(* IEC 61131-3 sources: Test-Git_ESME26/TestProgettoESME_26.fbsproj/PacDriveLib Migration/Motion/Control, 3 files *)

(* ---- PDL_FB_Brake.fb.st ---- *)
FUNCTION_BLOCK PDL_FB_Brake
VAR_INPUT
	i_xEnable  : BOOL;
	i_xRelease : BOOL;
	i_ifDrive  : Moin.IF_Axis;
END_VAR
VAR_OUTPUT
	q_xActive   : BOOL;
	q_xReady    : BOOL;
	q_etDiag    : GD.ET_Diag     := GD.ET_Diag.Ok;
	q_etDiagExt : PDL_ET_DiagExt := PDL_ET_DiagExt.Disabled;
	q_sMsg      : STRING[80];
	q_xReleased : BOOL;
END_VAR
VAR
	xSuccess                 : BOOL;
	ifDeviceTreeObjectAccess : UFMPLCI.IF_DeviceTreeObjectAccess;
	sDriveName               : STRING(80);
	ifBrakeAccess            : DDI.IF_BrakeAccess;
	ifBrake                  : DDI.IF_Brake;
	ifGetParentDevice        : DTSI.IF_GetParentDevice;
	ifDeviceAccess           : DTSI.IF_DeviceAccess;
	ifWorkingModeAccess      : CFDI.IF_WorkingModeAccess;
	ifWorkingMode            : CFDI.IF_WorkingMode;
	etWorkingState           : CFDI.ET_WorkingState;
	etSercosState            : SMI.ET_SercosState;
	etAxisState              : MOIN.ET_AxisState;
	etDiagExt                : PDL_ET_DiagExt := PDL_ET_DiagExt.Disabled;
	diState                  : DINT;
	xEnableFlag              : BOOL;
	fbLoggerPoint            : APL.FB_LoggerPoint;
	fbBrakeReleaseSet        : FB_BrakeReleaseSet;
	fbBrakeDisconnectionTime : FB_BrakeDisconnectionTime;
	fbBrakeCouplingTime      : FB_BrakeCouplingTime;
	xError                   : BOOL;
	tonTimeOutBrake          : Standard.TON;
	tonTimeOutException      : Standard.TON;
	tBrakeCouplingTemp       : TIME := T#500MS;
	tBrakeDisconnectTemp     : TIME := T#500MS;
	sResultMsg               : STRING(80);
	etResult                 : SE_Async.ET_Result;

END_VAR
VAR CONSTANT
	c_timTimeOutException : TIME := T#1S;
END_VAR

IF i_xEnable AND NOT xEnableFlag THEN (* Input action *)
	xEnableFlag := TRUE;

	THIS^.fbLoggerPoint.AddLogEntry(
		i_etLogLevel := APL.ET_LogLevel.UserAction,
		i_etDiag     := q_etDiag,
		i_udiDiagExt := q_etDiagExt,
		i_sMessage   := 'enable function block',
		q_etDiag     =>,
		q_etDiagExt  => );

	q_xActive   := TRUE;
	q_xReady    := FALSE;
	q_xReleased := FALSE;
	SetDiagOutput(
		i_etDiag    := GD.ET_Diag.Ok,
		i_etDiagExt := PDL_ET_DiagExt.Initializing,
		i_sMsg      := '');
	xSuccess := InitInterfaces();
	IF NOT xSuccess THEN
		RETURN;
	ELSE
		IF SE_Async.G_ifAsyncMgr.xInitDone THEN
			q_xReady    := TRUE;
			q_xReleased := (ifBrake.BrakeState = DDI.ET_BrakeState.released);
			IF q_xReleased THEN // Bremse is open --> wait for closing Brake (i_xRelease = false)
				SetDiagOutput(
					i_etDiag    := GD.ET_Diag.Ok,
					i_etDiagExt := PDL_ET_DiagExt.WaitForNotRelease,
					i_sMsg      := '');
				diState := 40;
			ELSE // brake is closed --> wait for opening brake (i_xRelease = true)
				SetDiagOutput(
					i_etDiag    := GD.ET_Diag.Ok,
					i_etDiagExt := PDL_ET_DiagExt.WaitForRelease,
					i_sMsg      := '');
				diState := 10;
			END_IF
		ELSE
			SE_Async.G_ifAsyncMgr.Init();
			diState := 150;
		END_IF
	END_IF

ELSIF NOT i_xEnable AND xEnableFlag AND q_xActive THEN
	xEnableFlag := FALSE;
	THIS^.fbLoggerPoint.AddLogEntry(
		i_etLogLevel := APL.ET_LogLevel.UserAction,
		i_etDiag     := q_etDiag,
		i_udiDiagExt := q_etDiagExt,
		i_sMessage   := 'disable function block',
		q_etDiag     =>,
		q_etDiagExt  => );
	SetDiagOutput(
		i_etDiag    := GD.ET_Diag.Ok,
		i_etDiagExt := PDL_ET_DiagExt.WaitUntilDisabled,
		i_sMsg      := '');

	q_xReady := FALSE;
	IF diState = 10 THEN // Brake is already closed
		diState := 120;
	ELSE
		fbBrakeReleaseSet.ifBrake  := ifBrake;
		fbBrakeReleaseSet.xRelease := FALSE;
		SE_Async.G_ifAsyncMgr.Start(
			i_ifAsync    := fbBrakeReleaseSet,
			q_etResult   => etResult,
			q_sResultMsg => sResultMsg,
			q_xError     => xError);
		IF xError THEN
			diState := 120;
		ELSE
			tonTimeOutBrake(IN := FALSE, PT := c_timTimeOutException);
			diState := 100;
		END_IF
	END_IF
END_IF

IF q_xReady THEN
	etSercosState  := FC_GetSercosState();
	etWorkingState := ifWorkingMode.ActualState;
	etAxisState    := i_ifDrive.etAxisState;
	IF etSercosState <> SMI.ET_SercosState.Phase4 THEN
		q_xReady    := FALSE;
		q_xReleased := FALSE;
		SetDiagOutput(
			i_etDiag    := GD.ET_Diag.SercosConditionInvalid,
			i_etDiagExt := PDL_ET_DiagExt.SercosNotInPhaseFour,
			i_sMsg      := 'Sercos not in phase four');
		diState := 0;
	ELSIF etWorkingState = CFDI.ET_WorkingState.Deactivated THEN
		q_xReady    := FALSE;
		q_xReleased := FALSE;
		SetDiagOutput(
			i_etDiag    := GD.ET_Diag.DriveConditionInvalid,
			i_etDiagExt := PDL_ET_DiagExt.DriveNotReady,
			i_sMsg		:= STANDARD.CONCAT(sDriveName, '.WorkingMode = deactivated'));
		diState := 0;
	ELSIF etAxisState <> Moin.ET_AxisState.Disabled THEN
		q_xReady    := FALSE;
		q_xReleased := FALSE;
		SetDiagOutput(
			i_etDiag    := GD.ET_Diag.DriveConditionInvalid,
			i_etDiagExt := PDL_ET_DiagExt.DriveNotReady,
			i_sMsg		:= STANDARD.CONCAT(sDriveName, '.AxisState <> Disabled; Drive has to be disabled'));
		diState := 0;
	END_IF
END_IF

CASE diState OF
	0: (* No operation / FB disabled *)
		;
	10: // Brake closed, wait for releasing Brake (i_xRelease = true)
		IF i_xRelease THEN // input release Brake
			fbLoggerPoint.AddLogEntry(
				i_etLogLevel := APL.ET_LogLevel.UserAction,
				i_etDiag     := q_etDiag,
				i_udiDiagExt := q_etDiagExt,
				i_sMessage   := 'Release Brake - read out disconnection time',
				q_etDiag     =>,
				q_etDiagExt  => );
			etSercosState := FC_GetSercosState();
			fbBrakeDisconnectionTime.ifBrake  := ifBrake;
			SE_Async.G_ifAsyncMgr.Start(
				i_ifAsync    := fbBrakeDisconnectionTime, // read Disconnecting time from Drive
				q_etResult   => etResult,
				q_sResultMsg => sResultMsg,
				q_xError     => xError);
			IF xError THEN
				IF etResult = SE_Async.ET_Result.MaxNumOfReusableObjectsExceeded THEN
					diState := diState; // Try again to Start Async in next cycle
				ELSE
					AsyncExtDiagTranslation();
					diState := 200;
				END_IF
			ELSE
				tonTimeOutBrake(IN := FALSE, PT := c_timTimeOutException);
				diState := 15;
			END_IF
		END_IF
	15: // Wait for BrakeDisconnectionTime has been read
		tonTimeOutBrake(IN := TRUE);
		IF fbBrakeDisconnectionTime.xDone THEN
			tBrakeDisconnectTemp       := fbBrakeDisconnectionTime.timTime;
			fbBrakeReleaseSet.ifBrake  := ifBrake;
			fbBrakeReleaseSet.xRelease := TRUE;
			SE_Async.G_ifAsyncMgr.Start(
				i_ifAsync    := fbBrakeReleaseSet,
				q_etResult   => etResult,
				q_sResultMsg => sResultMsg,
				q_xError     => xError);
			IF xError THEN
				IF etResult = SE_Async.ET_Result.MaxNumOfReusableObjectsExceeded THEN
					diState := diState; // Try again to Start Async in next cycle
				ELSE
					AsyncExtDiagTranslation();
					diState := 200;
				END_IF
			ELSE
				fbLoggerPoint.AddLogEntry(
					i_etLogLevel := APL.ET_LogLevel.DebugMessage,
					i_etDiag     := q_etDiag,
					i_udiDiagExt := q_etDiagExt,
					i_sMessage   := 'Release Brake - brake release set',
					q_etDiag     =>,
					q_etDiagExt  => );
				tonTimeOutBrake(IN := FALSE, PT := c_timTimeOutException);
				diState := 20;
			END_IF
		ELSIF tonTimeOutBrake.Q THEN
			SetDiagOutput(
				i_etDiag    := GD.ET_Diag.UnexpectedProgramBehavior,
				i_etDiagExt := PDL_ET_DiagExt.AsyncAddWasNotSuccessful,
				i_sMsg      := 'Timeout at read of BrakeDisconnectionTime');
			diState := 200;
		END_IF
	20: // Wait for Brake is release, Release Commando Done
		tonTimeOutBrake(IN := TRUE);
		IF fbBrakeReleaseSet.xDone THEN
			SetDiagOutput(
				i_etDiag    := GD.ET_Diag.Ok,
				i_etDiagExt := PDL_ET_DiagExt.WaitUntilBrakeReleased,
				i_sMsg      := '');
			tonTimeOutBrake(IN := FALSE, PT := tBrakeDisconnectTemp);
			tonTimeOutException(IN := FALSE, PT := c_timTimeOutException);
			diState := 25;
		ELSIF tonTimeOutBrake.Q THEN
			SetDiagOutput(
				i_etDiag    := GD.ET_Diag.UnexpectedProgramBehavior,
				i_etDiagExt := PDL_ET_DiagExt.AsyncAddWasNotSuccessful,
				i_sMsg      := 'Timeout at BrakeReleaseSet');
			diState := 200;
		END_IF
	25: // wait till brake has to be open (check both, system signal and own time out)
		tonTimeOutBrake(IN := TRUE);
		tonTimeOutException(IN := TRUE);
		IF tonTimeOutBrake.Q THEN
			IF (ifBrake.BrakeState = DDI.ET_BrakeState.released) THEN // Brake is released
				q_xReleased := TRUE;
				SetDiagOutput(
					i_etDiag    := GD.ET_Diag.Ok,
					i_etDiagExt := PDL_ET_DiagExt.WaitForNotRelease,
					i_sMsg      := '');
				diState := 40;
			ELSE
				SetDiagOutput(
					i_etDiag    := GD.ET_Diag.UnexpectedProgramBehavior,
					i_etDiagExt := PDL_ET_DiagExt.BrakeStateChangedNotInTime,
					i_sMsg      := 'Timeout at wait for Brake Release');
				diState := 200;
			END_IF
		ELSIF tonTimeOutException.Q THEN
			SetDiagOutput(
				i_etDiag    := GD.ET_Diag.UnexpectedProgramBehavior,
				i_etDiagExt := PDL_ET_DiagExt.BrakeStateChangedNotInTime,
				i_sMsg      := 'Timeout at wait for Brake Release');
			diState := 200;
		END_IF
	40: // Brake released, wait for Brake is coupled (i_xRelease = FALSE)
		IF NOT i_xRelease THEN
			fbLoggerPoint.AddLogEntry(
				i_etLogLevel := APL.ET_LogLevel.UserAction,
				i_etDiag     := q_etDiag,
				i_udiDiagExt := q_etDiagExt,
				i_sMessage   := 'Close Brake - read out coupling time',
				q_etDiag     =>,
				q_etDiagExt  => );
			fbBrakeCouplingTime.ifBrake  := ifBrake;
			SE_Async.G_ifAsyncMgr.Start(
				i_ifAsync    := fbBrakeCouplingTime,
				q_etResult   => etResult,
				q_sResultMsg => sResultMsg,
				q_xError     => xError);
			IF xError THEN
				IF etResult = SE_Async.ET_Result.MaxNumOfReusableObjectsExceeded THEN
					diState := diState; // Try again to Start Async in next cycle
				ELSE
					AsyncExtDiagTranslation();
					diState := 200;
				END_IF
			ELSE
				tonTimeOutBrake(IN := FALSE, PT := c_timTimeOutException);
				diState := 45;
			END_IF
		END_IF
	45: // wait for BrakeCouplingTime has been read out
		tonTimeOutBrake(IN := TRUE);
		IF fbBrakeCouplingTime.xDone THEN
			tBrakeCouplingTemp         := fbBrakeCouplingTime.timTime;
			fbBrakeReleaseSet.ifBrake  := ifBrake;
			fbBrakeReleaseSet.xRelease := FALSE;
			SE_Async.G_ifAsyncMgr.Start(
				i_ifAsync    := fbBrakeReleaseSet,
				q_etResult   => etResult,
				q_sResultMsg => sResultMsg,
				q_xError     => xError);
			IF xError THEN
				AsyncExtDiagTranslation();
				diState := 200;
			ELSE
				fbLoggerPoint.AddLogEntry(
					i_etLogLevel := APL.ET_LogLevel.DebugMessage,
					i_etDiag     := q_etDiag,
					i_udiDiagExt := q_etDiagExt,
					i_sMessage   := 'Close Brake - brake release set',
					q_etDiag     =>,
					q_etDiagExt  => );
				tonTimeOutBrake(IN := FALSE, PT := c_timTimeOutException);
				diState := 50;
			END_IF
		ELSIF tonTimeOutBrake.Q THEN
			SetDiagOutput(
				i_etDiag    := GD.ET_Diag.UnexpectedProgramBehavior,
				i_etDiagExt := PDL_ET_DiagExt.AsyncAddWasNotSuccessful,
				i_sMsg      := 'Timeout at read of BrakeCouplingTime');
			diState := 200;
		END_IF
	50: // Wait for BrakeRelaseSet Done
		tonTimeOutBrake(IN := TRUE);
		IF fbBrakeReleaseSet.xDone THEN
			SetDiagOutput(
				i_etDiag    := GD.ET_Diag.Ok,
				i_etDiagExt := PDL_ET_DiagExt.WaitUntilBrakeClosed,
				i_sMsg      := '');
			tonTimeOutBrake(IN := FALSE, PT := tBrakeCouplingTemp);
			tonTimeOutException(IN := FALSE, PT := c_timTimeOutException);
			diState := 55;
		ELSIF tonTimeOutBrake.Q THEN
			SetDiagOutput(
				i_etDiag    := GD.ET_Diag.UnexpectedProgramBehavior,
				i_etDiagExt := PDL_ET_DiagExt.AsyncAddWasNotSuccessful,
				i_sMsg      := 'Timeout at BrakeReleaseSet');
			diState := 200;
		END_IF
	55: // wait till brake is closed (check both, system signal and own time out)
		tonTimeOutBrake(IN := TRUE);
		tonTimeOutException(IN := TRUE);
		IF tonTimeOutBrake.Q THEN
			IF (ifBrake.BrakeState = DDI.ET_BrakeState.coupled)  THEN
				tonTimeOutException(IN := FALSE);
				tonTimeOutBrake(IN := FALSE);
				q_xReleased := FALSE;
				SetDiagOutput(
					i_etDiag    := GD.ET_Diag.Ok,
					i_etDiagExt := PDL_ET_DiagExt.WaitForRelease,
					i_sMsg      := '');
				diState := 10;
			ELSE
				SetDiagOutput(
					i_etDiag    := GD.ET_Diag.UnexpectedProgramBehavior,
					i_etDiagExt := PDL_ET_DiagExt.BrakeStateChangedNotInTime,
					i_sMsg      := 'Timeout at wait for Brake coupled');
				diState := 200;
			END_IF
		ELSIF tonTimeOutBrake.Q THEN
			SetDiagOutput(
				i_etDiag    := GD.ET_Diag.UnexpectedProgramBehavior,
				i_etDiagExt := PDL_ET_DiagExt.BrakeStateChangedNotInTime,
				i_sMsg      := 'Timeout at wait for Brake Close');
			diState := 200;
		END_IF

		//---------------------------------------------------------------------------------
	100:
		tonTimeOutBrake(IN := TRUE);
		IF fbBrakeReleaseSet.xDone THEN
			IF i_ifDrive.etAxisState = MOIN.ET_AxisState.Disabled THEN
				tonTimeOutBrake(IN := FALSE, PT := c_timTimeOutException);
				diState := 110;
			ELSE
				diState := 120;
			END_IF
		ELSIF tonTimeOutBrake.Q THEN
			SetDiagOutput(
				i_etDiag    := GD.ET_Diag.UnexpectedProgramBehavior,
				i_etDiagExt := PDL_ET_DiagExt.AsyncAddWasNotSuccessful,
				i_sMsg      := 'Timeout at FC_BrakeReleaseSet');
			diState := 120;
		END_IF
	110: (* AxisState = 1 or 2 *)
		tonTimeOutBrake(IN := TRUE);
		IF (ifBrake.BrakeState = DDI.ET_BrakeState.coupled) THEN
			tonTimeOutBrake(IN := FALSE, PT := tBrakeCouplingTemp);
			diState := 115;
		ELSIF tonTimeOutBrake.Q THEN
			SetDiagOutput(
				i_etDiag    := GD.ET_Diag.UnexpectedProgramBehavior,
				i_etDiagExt := PDL_ET_DiagExt.BrakeStateChangedNotInTime,
				i_sMsg      := 'Timeout at wait for Brake Close');
			diState := 120;
		END_IF
	115:
		tonTimeOutBrake(IN := TRUE);
		IF tonTimeOutBrake.Q THEN
			diState := 120;
		END_IF
	120:
		q_xActive   := FALSE;
		q_xReady    := FALSE;
		q_xReleased := FALSE;
		SetDiagOutput(
			i_etDiag    := GD.ET_Diag.Ok,
			i_etDiagExt := PDL_ET_DiagExt.Disabled,
			i_sMsg      := '');
		tonTimeOutBrake(IN := FALSE);
		diState := 0;

	150:
		SE_Async.G_ifAsyncMgr.Init(
			q_xError     => xError,
			q_etResult   => etResult,
			q_sResultMsg => sResultMsg);
		IF xError THEN
			AsyncExtDiagTranslation();
			diState := 200;
		ELSIF SE_Async.G_ifAsyncMgr.xInitDone THEN
			q_xReady    := TRUE;
			q_xReleased := (ifBrake.BrakeState = DDI.ET_BrakeState.released);
			IF q_xReleased THEN // Bremse is open --> wait for closing Brake (i_xRelease = false)
				SetDiagOutput(
					i_etDiag    := GD.ET_Diag.Ok,
					i_etDiagExt := PDL_ET_DiagExt.WaitForNotRelease,
					i_sMsg      := '');
				diState := 40;
			ELSE // brake is closed --> wait for opening brake (i_xRelease = true)
				SetDiagOutput(
					i_etDiag    := GD.ET_Diag.Ok,
					i_etDiagExt := PDL_ET_DiagExt.WaitForRelease,
					i_sMsg      := '');
				diState := 10;
			END_IF
		END_IF

	200:
		q_xReady    := FALSE;
		q_xReleased := (ifBrake.BrakeState = DDI.ET_BrakeState.released);
		diState := 0;

END_CASE

(* ---- PDL_FB_DriveEnable.fb.st ---- *)
FUNCTION_BLOCK PDL_FB_DriveEnable
VAR_INPUT
	i_xEnable      : BOOL; (* Enable of FB *)
	i_ifDrive      : MOIN.IF_Axis; (* Axis *)
	i_xEnableDrive : BOOL; (* Power on *)
	i_xDiagQuit    : BOOL; (* reset error *)
END_VAR

VAR_OUTPUT
	q_xActive       : BOOL; (* FB enabled*)
	q_xReady        : BOOL;
	q_etDiag        : GD.ET_Diag     := GD.ET_Diag.Ok;
	q_etDiagExt     : PDL_ET_DiagExt := PDL_ET_DiagExt.Disabled;
	q_sMsg          : STRING[80];
	q_xDriveEnabled : BOOL; (* power is on*)
END_VAR

VAR
	xInterfacesInitialised : BOOL;

	xEnableFlag : BOOL;
	diState     : DINT;

	rtrigDiagQuit    : Standard.R_TRIG;
	xDriveEnabledOld : BOOL;

	fbLoggerPoint : APL.FB_LoggerPoint;

	fbPower : PLCO.MC_Power;
	fbStop  : PLCO.MC_Stop;
	fbReset	: PLCO.MC_Reset;

	ifDeviceTreeObjectAccess      : UFMPLCI.IF_DeviceTreeObjectAccess;
	sDriveName                    : STRING(80);
	ifGetParentDevice             : DTSI.IF_GetParentDevice;
	ifDiagnostic                  : UFMPLCI.IF_Diagnostic;
	ifDiagnosticAccess            : UFMPLCI.IF_DiagnosticAccess;
	ifDeviceAccess                : DTSI.IF_DeviceAccess;
	ifPowerSupply                 : DDI.IF_PowerSupply;
	ifPowerSupplyAccess           : DDI.IF_PowerSupplyAccess;
	ifDrivePowerSupply            : DDI.IF_DrivePowerSupply;
	ifDrivePowerSupplyAccess      : DDI.IF_DrivePowerSupplyAccess;
	ifDriveConfigAccess           : DDI.IF_DriveConfigAccess;
	ifDriveConfig                 : DDI.IF_DriveConfig;
	ifWorkingModeAccess           : CFDI.IF_WorkingModeAccess;
	ifWorkingMode                 : CFDI.IF_WorkingMode;
	ifPowerSupplyDiagnosticAccess : UFMPLCI.IF_DiagnosticAccess;
	ifPowerSupplyDiagnostic       : UFMPLCI.IF_Diagnostic;
	ifPowerSupplyDevice           : DDI.DeviceTypeInterfaces.IF_Device_Type;
	xSuccess                      : BOOL;
	etSercosState                 : SMI.ET_SercosState;
	tonTimeOut                    : Standard.TON;
	xDriveIsReal                  : BOOL;
END_VAR
VAR CONSTANT
	c_timTimeoutPowerSupplyReady  : TIME := T#2000MS;
	c_timTimeoutPowerSupplyEnable : TIME := T#2000MS;
END_VAR

(*--------------------------------------------------------------------------------------------------------------------------------------------*)
//Enable
{region "enable"}
IF i_xEnable AND NOT xEnableFlag THEN
	xEnableFlag := TRUE;

	THIS^.fbLoggerPoint.AddLogEntry(	i_etLogLevel	:= APL.ET_LogLevel.UserAction,
										i_etDiag		:= q_etDiag,
										i_udiDiagExt	:= q_etDiagExt,
										i_sMessage		:= 'enable function block',
										q_etDiag		=> ,
										q_etDiagExt		=> );
	q_xActive			:= TRUE;
	q_xDriveEnabled		:= FALSE;

	IF NOT Init() THEN
		q_xReady			    := FALSE;
		xInterfacesInitialised  := FALSE;
		diState := 200;
	ELSE
		q_xReady 				:= TRUE;
		xInterfacesInitialised  := TRUE;
		SetDiagOutput(	i_etDiag	:= GD.ET_Diag.Ok,
						i_etDiagExt := PDL_ET_DiagExt.WaitForEnableDrive,
						i_sMsg		:= '');
		diState	:= 10;
	END_IF
{endregion}

(*--------------------------------------------------------------------------------------------------------------------------------------------*)
//Disable
{region "disable"}
ELSIF NOT i_xEnable AND xEnableFlag THEN
	xEnableFlag := FALSE;
	THIS^.fbLoggerPoint.AddLogEntry(	i_etLogLevel	:= APL.ET_LogLevel.UserAction,
										i_etDiag		:= q_etDiag,
										i_udiDiagExt	:= q_etDiagExt,
										i_sMessage		:= 'disable function block',
										q_etDiag		=> ,
										q_etDiagExt		=> );
	q_xReady			:= FALSE;
	IF xInterfacesInitialised THEN
		SetDiagOutput(	i_etDiag	:= GD.ET_Diag.Ok,
						i_etDiagExt := PDL_ET_DiagExt.WaitUntilDriveDisabled,
						i_sMsg		:= '');

		diState := 100; // whait till axis disabled
	ELSE
		q_xActive			:= FALSE;
		q_xDriveEnabled		:= FALSE;

		SetDiagOutput(	i_etDiag	:= GD.ET_Diag.Ok,
						i_etDiagExt := PDL_ET_DiagExt.Disabled,
						i_sMsg		:= '');
		diState	:= 0;
	END_IF
END_IF
{endregion}

(*--------------------------------------------------------------------------------------------------------------------------------------------*)
// Cyclic when enabled
{region "cyclic"}
IF xInterfacesInitialised AND q_xActive THEN
	q_xDriveEnabled :=  i_ifDrive.etAxisState >= MOIN.ET_AxisState.Standstill;
	etSercosState := FC_GetSercosState();
	fbReset( Execute := FALSE );

	IF xDriveIsReal AND_THEN ifPowerSupplyDiagnostic.DiagClass >= 3 THEN
		fbPower( Enable := FALSE );
		q_xReady	:= FALSE;
		SetDiagOutput(	i_etDiag	:= GD.ET_Diag.PowerSupplyConditionInvalid,
						i_etDiagExt := PDL_ET_DiagExt.PowerSupplyNotReady,
						i_sMsg		:= SE_CTBX.FC_MultiConcat(	i_sString1 := 'DiagCode: ',
														i_sString2 := TO_STRING(ifPowerSupplyDiagnostic.DiagCode),
														i_sString3 := ' - DiagMsg: ',
														i_sString4 := ifPowerSupplyDiagnostic.DiagMsg));
		diState := 200;

	//check for drive errors
	ELSIF ifDiagnostic.DiagClass >= 3 THEN
		fbPower( Enable := FALSE );
		q_xReady		:= FALSE;
		q_xDriveEnabled := FALSE;
		SetDiagOutput(	i_etDiag	:= GD.ET_Diag.DriveConditionInvalid,
						i_etDiagExt := PDL_ET_DiagExt.DriveNotReady,
						i_sMsg		:= SE_CTBX.FC_MultiConcat(	i_sString1 := 'DiagCode: ',
																i_sString2 := TO_STRING(ifDiagnostic.DiagCode),
																i_sString3 := ' - DiagMsg: ',
																i_sString4 := ifDiagnostic.DiagMsg));
		diState := 200;

	//check sercos state
	ELSIF etSercosState <> SMI.ET_SercosState.Phase4 THEN
		fbPower( Enable := FALSE );
		q_xReady:= FALSE;
		q_xDriveEnabled:= FALSE;
		SetDiagOutput(	i_etDiag	:= GD.ET_Diag.SercosConditionInvalid,
						i_etDiagExt := PDL_ET_DiagExt.SercosNotInPhaseFour,
						i_sMsg		:= 'Sercos not in phase four');
		diState:= 200;

	//check inverter enable
	ELSIF xDriveIsReal AND_THEN NOT ifDrivePowerSupply.InverterEnable AND i_xEnableDrive THEN
		fbPower( Enable := FALSE );
		q_xReady			:= FALSE;
		q_xDriveEnabled		:= FALSE;
		SetDiagOutput(	i_etDiag	:= GD.ET_Diag.DriveConditionInvalid,
						i_etDiagExt := PDL_ET_DiagExt.InverterEnableOff,
						i_sMsg		:= sDriveName);
		diState := 200;
	END_IF

	//stop/disable drive
	IF    NOT i_xEnableDrive
	  AND diState = 10
	  AND fbPower.Enable
	THEN
		THIS^.fbLoggerPoint.AddLogEntry(	i_etLogLevel	:= APL.ET_LogLevel.UserAction,
											i_etDiag		:= q_etDiag,
											i_udiDiagExt	:= q_etDiagExt,
											i_sMessage		:= 'disable drive',
											q_etDiag		=> ,
											q_etDiagExt		=> );

		SetDiagOutput(	i_etDiag	:= GD.ET_Diag.Ok,
						i_etDiagExt := PDL_ET_DiagExt.WaitUntilDriveDisabled,
						i_sMsg		:= '');

		//if power on -> stop first
		IF fbPower.Status THEN
			diState := 30;
		ELSE
			diState := 100;
		END_IF
	END_IF

END_IF

IF q_xActive THEN
	rtrigDiagQuit(CLK := i_xDiagQuit);
END_IF
{endregion}

(*--------------------------------------------------------------------------------------------------------------------------------------------*)
//state machine
CASE diState OF

(*********************************************************************************************************************)
	0:	//Error or Not Enabled
		;

(*********************************************************************************************************************)
	10:	//enable drive
{region "enableDrive"}
		fbStop(Axis := i_ifDrive, Execute := FALSE );

		//set diag outpupt after enable cmd
		IF 	  i_xEnableDrive
		  AND NOT fbPower.Enable
		  AND i_xEnable
		THEN
			IF xDriveIsReal AND_THEN NOT ifPowerSupply.PowerSupplyCheck THEN
				ifPowerSupply.PowerSupplyCheckSet	:= TRUE;
				SetDiagOutput(	i_etDiag	:= GD.ET_Diag.Ok,
								i_etDiagExt := PDL_ET_DiagExt.WaitUntilPowerSupplyReady,
								i_sMsg		:= '');
				tonTimeout(IN := FALSE, PT := c_timTimeoutPowerSupplyReady);		(* init Timeout for PS Ready *)
				diState	:= 20;
				RETURN;
			ELSE
				THIS^.fbLoggerPoint.AddLogEntry(	i_etLogLevel	:= APL.ET_LogLevel.UserAction,
													i_etDiag		:= q_etDiag,
													i_udiDiagExt	:= q_etDiagExt,
													i_sMessage		:= 'enable drive',
													q_etDiag		=> ,
													q_etDiagExt		=> );

				SetDiagOutput(	i_etDiag	:= GD.ET_Diag.Ok,
								i_etDiagExt := PDL_ET_DiagExt.WaitUntilDriveEnabled,
								i_sMsg		:= '');
			END_IF
		END_IF

		//cmd power on
		fbPower( Enable :=  i_xEnableDrive AND i_xEnable );
		q_xDriveEnabled :=  i_ifDrive.etAxisState >= MOIN.ET_AxisState.Standstill;

		//set diag output when on
		IF    q_xDriveEnabled
		  AND NOT xDriveEnabledOld
		THEN
			SetDiagOutput(	i_etDiag	:= GD.ET_Diag.Ok,
							i_etDiagExt := PDL_ET_DiagExt.DriveEnabled,
							i_sMsg		:= '');
		END_IF

		//error
		IF fbPower.Error THEN
			q_xReady		:= FALSE;
			q_xDriveEnabled	:= FALSE;

			SetDiagOutput(	i_etDiag	:= GD.ET_Diag.UnexpectedProgramBehavior,
							i_etDiagExt := PDL_ET_DiagExt.UnexpectedFeedback,
							i_sMsg		:= CONCAT('MC_Power.ErrorID: ', PLCO.FC_EtResultToString( fbPower.ErrorID ) ));

			fbPower( Enable := FALSE );
			diState	:= 200;
		END_IF
{endregion}

(*********************************************************************************************************************)
	20: (* Wait for PowerSupply GroupState >= 2 *)
{region "error"}
		tonTimeout(IN := TRUE);
		IF ifPowerSupply.GroupState >= 2  THEN								(* GroupState on PS *)
			tonTimeout(IN := FALSE, PT := c_timTimeoutPowerSupplyEnable);	(* init Timeout for PS Enabled *)
			diState := 10;

		ELSIF tonTimeout.Q THEN
			q_xReady	:= FALSE;
			SetDiagOutput(	i_etDiag	:= GD.ET_Diag.PowerSupplyConditionInvalid,
							i_etDiagExt := PDL_ET_DiagExt.PowerSupplyNotReady,
							i_sMsg		:= SE_CTBX.FC_MultiConcat(	i_sString1 := 'DiagCode: ',
																	i_sString2 := TO_STRING(ifPowerSupplyDiagnostic.DiagCode),
																	i_sString3 := ' - DiagMsg: ',
																	i_sString4 := ifPowerSupplyDiagnostic.DiagMsg));
			diState := 10;
		END_IF
{endregion}

(*********************************************************************************************************************)
	30: //controllerStop
{region "controllerStop"}
		IF 	  i_ifDrive.etAxisState <> MOIN.ET_AxisState.Disabled
		  AND i_ifDrive.etAxisState <> MOIN.ET_AxisState.ErrorStop
		  AND i_ifDrive.etAxisState <> MOIN.ET_AxisState.Standstill
		  AND i_ifDrive.etAxisState <> MOIN.ET_AxisState.Stopping
		THEN
			fbStop.Execute 			:= TRUE;
			fbStop.Deceleration 	:= i_ifDrive.lrErrorStopDec;
			fbStop.Jerk 			:= i_ifDrive.lrErrorStopJerk;
		END_IF

		fbStop();

		//stopping done
		IF 	  i_ifDrive.etAxisState = MOIN.ET_AxisState.Disabled
		  OR  i_ifDrive.etAxisState = MOIN.ET_AxisState.ErrorStop
		  OR  i_ifDrive.etAxisState = MOIN.ET_AxisState.Standstill
		  OR  fbStop.Done
		THEN
			fbStop( Axis := i_ifDrive, Execute := FALSE );

			diState := 100;
		END_IF

		//error
		IF fbStop.Error AND fbStop.ErrorId <> PLCO.ET_Result.StoppingInterrupted THEN
			q_xReady		:= FALSE;
			q_xDriveEnabled	:= FALSE;

			fbStop( Axis := i_ifDrive, Execute := FALSE );
			SetDiagOutput(	i_etDiag	:= GD.ET_Diag.UnexpectedProgramBehavior,
							i_etDiagExt := PDL_ET_DiagExt.UnexpectedFeedback,
							i_sMsg		:= CONCAT('MC_Stop.ErrorID: ', PLCO.FC_EtResultToString(fbStop.ErrorID) ));
			diState := 100;
		END_IF
{endregion}

(*********************************************************************************************************************)
	100: //disable drive
{region "disableDrive"}
		fbStop( Execute := FALSE );
		fbPower( Enable :=  FALSE );

		q_xDriveEnabled := i_ifDrive.etAxisState >= MOIN.ET_AxisState.Standstill;

		//wait for power off
		IF NOT q_xDriveEnabled THEN
			IF NOT i_xEnable THEN
				q_xActive := FALSE;
				SetDiagOutput(	i_etDiag	:= GD.ET_Diag.Ok,
								i_etDiagExt := PDL_ET_DiagExt.Disabled,
								i_sMsg		:= '');
				diState	:= 0;
			ELSE
				SetDiagOutput(	i_etDiag	:= GD.ET_Diag.Ok,
								i_etDiagExt := PDL_ET_DiagExt.WaitForEnableDrive,
								i_sMsg		:= '');
				diState	:= 10;
			END_IF
		END_IF

		//error
		IF fbPower.Error THEN
			q_xReady		:= FALSE;
			q_xDriveEnabled	:= FALSE;

			SetDiagOutput(	i_etDiag	:= GD.ET_Diag.UnexpectedProgramBehavior,
							i_etDiagExt := PDL_ET_DiagExt.UnexpectedFeedback,
							i_sMsg		:= CONCAT('MC_Power.ErrorID: ', PLCO.FC_EtResultToString( fbPower.ErrorID ) ));
			fbStop( Execute := FALSE );
		  	IF i_xEnable THEN
				diState	:= 200;
			ELSE
				diState	:= 0;
			END_IF
		END_IF
{endregion}

(*********************************************************************************************************************)
	200: //error
{region "error"}
		IF rtrigDiagQuit.Q //wait for cmd diag quit
		THEN
			THIS^.fbLoggerPoint.AddLogEntry(	i_etLogLevel	:= APL.ET_LogLevel.UserAction,
												i_etDiag		:= q_etDiag,
												i_udiDiagExt	:= q_etDiagExt,
												i_sMessage		:= 'diag quit',
												q_etDiag		=> ,
												q_etDiagExt		=> );
			IF NOT Init() THEN
				// error was not quittable -> keep error state
				xInterfacesInitialised := FALSE;

			ELSE
				// reset error
				IF i_ifDrive.etAxisState = MOIN.ET_AxisState.ErrorStop THEN
					fbReset( Execute := TRUE );
				END_IF

				xInterfacesInitialised := TRUE;
				q_xReady := TRUE;
				q_etDiag := GD.ET_Diag.Ok; // has to be done outside of SetDiagOutput too, because new Diagnosis is only set if FB does not signal Error
				SetDiagOutput(	i_etDiag	:= GD.ET_Diag.Ok,
								i_etDiagExt := PDL_ET_DiagExt.WaitForEnableDrive,
								i_sMsg		:= '');
				diState := 10;
			END_IF
		END_IF
{endregion}

END_CASE
(*--------------------------------------------------------------------------------------------------------------------------------------------*)
xDriveEnabledOld := q_xDriveEnabled;

(* ---- PDL_FB_YOffsetCorrection.fb.st ---- *)
{attribute 'no_assign'}
FUNCTION_BLOCK PDL_FB_YOffsetCorrection

VAR_INPUT
	i_xEnable				: BOOL;								(* Enables the FB *)
	i_ifDrive				: MOIN.IF_Axis;						(* Slave Axis *)
	i_lencMaster			: MOIN.IF_LogicalEncoder;			(* Master *)
	i_xStart				: BOOL;								(* Starts Correction *)
	i_lrCorrection			: LREAL;							(* Value of Correction *)
	i_lrXStartPos			: LREAL;							(* Start position of correction *)
	i_lrXFactor				: LREAL;							(* Distance covered by the master within which the correction is to be executed *)
	i_lrMaxCorrVel			: LREAL;							(* max velocity for correction *)
	i_lrMaxCorrAcc			: LREAL;							(* max acc/dec for correction *)
END_VAR

VAR_OUTPUT
	q_xActive				: BOOL;
	q_xReady				: BOOL;
	q_xCorrectionActive		: BOOL;
	q_etDiag				: GD.ET_Diag := GD.ET_Diag.OK;
	q_etDiagExt				: PDL_ET_DiagExt := PDL_ET_DiagExt.Disabled;
	q_sMsg					: STRING[80];
END_VAR

VAR
	xEnableFlag				: BOOL;
	diState					: DINT;
	xInterfacesInitialised	: BOOL;

	lrCorrVel				: LREAL;
	lrCorrAcc				: LREAL;
	lrCorrTime				: LREAL;
	diResult				: DINT;

	//superimposed movement
	fbMoveSuperimposed		: PLCO.MC_MoveSuperimposed;
	fbHalt					: PLCO.MC_Halt;

	//channels
	fbReadAxisInfo			: PLCO.MC_ReadAxisInfo;
	fbMultiComb				: MLTCMB.FB_MultiCombine<2>;
	fbPowerControlAxis		: PLCO.MC_Power;
	fbPowerOffsetAxis		: PLCO.MC_Power;
	fbSetPos				: PLCO.MC_SetPosition;
	ifControlChannel		: MOIN.IF_Axis;
	ifOffsetChannel			: MOIN.IF_Axis;
END_VAR

(*--------------------------------------------------------------------------------------------------------------------------------------------*)
//enable
{region "enable"}
IF i_xEnable AND NOT xEnableFlag THEN
	xEnableFlag := TRUE;

	q_xActive			:= TRUE;
	q_xReady			:= FALSE;
	q_xCorrectionActive := FALSE;

	SetDiagOutput(	i_etDiag	:= GD.ET_Diag.OK,
					i_etDiagExt := PDL_ET_DiagExt.Initializing,
					i_sMsg		:= '');

	xInterfacesInitialised := Init();
	IF NOT xInterfacesInitialised THEN
		RETURN;
	END_IF

	//set control channel to axis pos
	fbSetPos( Execute := FALSE );
	fbSetPos(	Axis		:= fbMultiComb.Channels[0],
				Execute		:= TRUE,
				Relative	:= FALSE,
				Position	:= i_ifDrive.lrPosition);

	IF fbSetPos.Error THEN
		SetDiagOutput(	i_etDiag	:= GD.ET_Diag.UnexpectedProgramBehavior,
						i_etDiagExt := PDL_ET_DiagExt.UnexpectedFeedback,
						i_sMsg		:= CONCAT('MC_SetPosition.ErrorId: ', PLCO.FC_EtResultToString(fbSetPos.ErrorId) ) );
		fbSetPos( Execute := FALSE );
		diState := 0;
		RETURN;
	END_IF

	//set offset to 0
	fbSetPos( Execute := FALSE );
	fbSetPos(	Axis		:= fbMultiComb.Channels[1],
				Execute		:= TRUE,
				Relative	:= FALSE,
				Position	:= 0);

	IF fbSetPos.Error THEN
		SetDiagOutput(	i_etDiag	:= GD.ET_Diag.UnexpectedProgramBehavior,
						i_etDiagExt := PDL_ET_DiagExt.UnexpectedFeedback,
						i_sMsg		:= CONCAT('MC_SetPosition.ErrorId: ', PLCO.FC_EtResultToString(fbSetPos.ErrorId) ) );
		fbSetPos( Execute := FALSE );
		diState := 0;
		RETURN;
	END_IF

	q_xReady := TRUE;

	SetDiagOutput(	i_etDiag	:= GD.ET_Diag.Ok,
					i_etDiagExt := PDL_ET_DiagExt.WaitForStart,
					i_sMsg		:= '');
	diState	:= 10;
{endregion}

(*--------------------------------------------------------------------------------------------------------------------------------------------*)
//disable
{region "disable"}
ELSIF NOT i_xEnable AND xEnableFlag THEN
	xEnableFlag := FALSE;
	xInterfacesInitialised := FALSE;

	q_xCorrectionActive					:= FALSE;
	q_xActive							:= FALSE;
	q_xReady							:= FALSE;

	//set axis relative
	fbSetPos( Execute := FALSE );
	fbSetPos(	Axis		:= i_ifDrive,
				Execute		:= TRUE,
				Relative	:= TRUE,
				Position	:= -fbMultiComb.Channels[1].lrPosition );

	IF fbSetPos.Error THEN
		SetDiagOutput(	i_etDiag	:= GD.ET_Diag.UnexpectedProgramBehavior,
						i_etDiagExt := PDL_ET_DiagExt.UnexpectedFeedback,
						i_sMsg		:= CONCAT('MC_SetPosition.ErrorId: ', PLCO.FC_EtResultToString(fbSetPos.ErrorId) ) );
		fbSetPos( Execute := FALSE );
		diState := 0;
		RETURN;
	END_IF

	//set offset to 0
	fbSetPos( Execute := FALSE );
	fbSetPos(	Axis		:= fbMultiComb.Channels[1],
				Execute		:= TRUE,
				Relative	:= FALSE,
				Position	:= 0);

	IF fbSetPos.Error THEN
		SetDiagOutput(	i_etDiag	:= GD.ET_Diag.UnexpectedProgramBehavior,
						i_etDiagExt := PDL_ET_DiagExt.UnexpectedFeedback,
						i_sMsg		:= CONCAT('MC_SetPosition.ErrorId: ', PLCO.FC_EtResultToString(fbSetPos.ErrorId) ) );
		fbSetPos( Execute := FALSE );
		diState := 0;
		RETURN;
	END_IF

	SetDiagOutput(	i_etDiag	:= GD.ET_Diag.Ok,
					i_etDiagExt := PDL_ET_DiagExt.Disabled,
					i_sMsg		:= '');
	diState := 0;
END_IF
{endregion}

(*--------------------------------------------------------------------------------------------------------------------------------------------*)
// Cyclic
{region "cyclic"}
IF i_ifDrive <> 0 THEN

	//read power on state...
	fbReadAxisInfo( Axis				:= i_ifDrive,
					Enable				:= TRUE);

	IF fbReadAxisInfo.Error THEN
		SetDiagOutput(	i_etDiag	:= GD.ET_Diag.UnexpectedProgramBehavior,
						i_etDiagExt := PDL_ET_DiagExt.UnexpectedFeedback,
						i_sMsg		:= CONCAT('MC_ReadAxisInfo.ErrorId: ', PLCO.FC_EtResultToString(fbReadAxisInfo.ErrorId) ) );
		fbReadAxisInfo( Enable := FALSE );
		fbMoveSuperimposed( Execute := FALSE );
		diState := 0;
	END_IF

	//... and switch on power at channels
	fbPowerControlAxis(	Axis   := fbMultiComb.Channels[0],
						Enable := fbReadAxisInfo.PowerOn);

	IF fbPowerControlAxis.Error THEN
		SetDiagOutput(	i_etDiag	:= GD.ET_Diag.UnexpectedProgramBehavior,
						i_etDiagExt := PDL_ET_DiagExt.UnexpectedFeedback,
						i_sMsg		:= CONCAT('MC_Power.ErrorId: ', PLCO.FC_EtResultToString(fbPowerControlAxis.ErrorId) ) );
		fbPowerControlAxis( Enable := FALSE );
		fbMoveSuperimposed( Execute := FALSE );
		diState := 0;
	END_IF

	fbPowerOffsetAxis(	Axis:= fbMultiComb.Channels[1],
						Enable:= fbReadAxisInfo.PowerOn);

	IF fbPowerOffsetAxis.Error THEN
		SetDiagOutput(	i_etDiag	:= GD.ET_Diag.UnexpectedProgramBehavior,
						i_etDiagExt := PDL_ET_DiagExt.UnexpectedFeedback,
						i_sMsg		:= CONCAT('MC_Power.ErrorId: ', PLCO.FC_EtResultToString(fbPowerOffsetAxis.ErrorId) ) );
		fbPowerOffsetAxis( Enable := FALSE );
		fbMoveSuperimposed( Execute := FALSE );
		diState := 0;
	END_IF

	//muticombine
	fbMultiComb(Slave			:= i_ifDrive,
				Execute			:=    fbReadAxisInfo.PowerOn
								  AND fbPowerControlAxis.Status
								  AND fbPowerOffsetAxis.Status
				);

	IF fbMultiComb.Error THEN
		SetDiagOutput(	i_etDiag	:= GD.ET_Diag.UnexpectedProgramBehavior,
						i_etDiagExt := PDL_ET_DiagExt.UnexpectedFeedback,
						i_sMsg		:= CONCAT('FB_MultiCombine.ErrorId: ', TO_STRING(fbMultiComb.ErrorId) ) );
		fbMultiComb( Execute := FALSE );
		fbMoveSuperimposed( Execute := FALSE );
		diState := 0;
	END_IF

ELSE
	SetDiagOutput(	i_etDiag	:= GD.ET_Diag.InputParameterInvalid,
					i_etDiagExt := PDL_ET_DiagExt.DriveInvalid,
					i_sMsg		:= 'i_ifDrive - Invalid Interface');
END_IF

ifControlChannel := fbMultiComb.Channels[0];
ifOffsetChannel  := fbMultiComb.Channels[1];
{endregion}

(*--------------------------------------------------------------------------------------------------------------------------------------------*)
// State machine
CASE diState OF

(*********************************************************************************************************************)
	0:	// error or disabled
		;

(*********************************************************************************************************************)
	10:	// Wait for Start
{region "waitForStartCmd"}
		IF i_xStart AND i_lencMaster.lrPosition < i_lrXStartPos THEN
			SetDiagOutput(	i_etDiag	:= GD.ET_Diag.Ok,
							i_etDiagExt := PDL_ET_DiagExt.WaitUntilMasterPositionGreaterXStartPosition,
							i_sMsg		:= '');

			diState	:= 20;
		END_IF

		//call fbHalt until finished (started in step 30)
		fbHalt(	Axis := ifOffsetChannel );
		IF fbHalt.Done THEN
			fbHalt( Execute := FALSE );
		END_IF

		IF fbHalt.Error THEN
			SetDiagOutput(	i_etDiag	:= GD.ET_Diag.UnexpectedProgramBehavior,
							i_etDiagExt := PDL_ET_DiagExt.UnexpectedFeedback,
							i_sMsg		:= CONCAT('MC_Halt.ErrorId: ', PLCO.FC_EtResultToString(fbHalt.ErrorId) ));
			fbHalt( Execute := FALSE );
			diState := 0;
			RETURN;
		END_IF

{endregion}

(*********************************************************************************************************************)
	20:	// wait  XPosition > XStart
{region "waitForStartPosition"}
		IF i_lencMaster.lrPosition >= i_lrXStartPos THEN
			lrCorrTime := ABS(i_lrXFactor / MAX(i_lencMaster.lrVelocity, 1.0));

			//calculate correction velocity
			lrCorrVel :=  ABS(i_lrCorrection / lrCorrTime * 1.5 );
			IF lrCorrVel > i_lrMaxCorrVel THEN
				lrCorrVel := i_lrMaxCorrVel;
			ELSIF lrCorrVel < i_lrMaxCorrVel / 1000.0 THEN
				lrCorrVel := i_lrMaxCorrVel / 1000.0;
			END_IF

			lrCorrAcc := lrCorrVel / lrCorrTime * 3.0;
			IF lrCorrAcc > i_lrMaxCorrAcc THEN
				lrCorrAcc := i_lrMaxCorrAcc;
			END_IF

			//start movement cmd...
			fbMoveSuperimposed( Execute := FALSE );
			fbMoveSuperimposed(	Axis			:= ifOffsetChannel,
								Execute			:= TRUE,
								Distance		:= i_lrCorrection,
								VelocityDiff	:= lrCorrVel,
								Acceleration	:= lrCorrAcc,
								Deceleration	:= lrCorrAcc );

			//...error
			IF fbMoveSuperimposed.Error THEN
				q_xCorrectionActive := FALSE;
				SetDiagOutput(	i_etDiag	:= GD.ET_Diag.UnexpectedProgramBehavior,
								i_etDiagExt := PDL_ET_DiagExt.UnexpectedFeedback,
								i_sMsg		:= CONCAT('MC_MoveSuperimposed.ErrorId: ', TO_STRING(fbMoveSuperimposed.ErrorId)));
				fbMoveSuperimposed( Execute := FALSE );
				diState := 0;

			ELSE
			//...success -> wait until finshed
				q_xCorrectionActive := TRUE;
				SetDiagOutput(	i_etDiag	:= GD.ET_Diag.Ok,
								i_etDiagExt := PDL_ET_DiagExt.WaitUntilYOffsetCorrectionFinished,
								i_sMsg		:= '');
				diState	:= 30;
			END_IF

		//user interrupt -> back to waiting
		ELSIF NOT i_xStart THEN
			q_xCorrectionActive := FALSE;

			SetDiagOutput(	i_etDiag	:= GD.ET_Diag.Ok,
							i_etDiagExt := PDL_ET_DiagExt.WaitForStart,
							i_sMsg		:= '');
			diState	:= 10;
		END_IF
{endregion}

(*********************************************************************************************************************)
	30:	// wait until finished
{region "waitUntilFinished"}
		fbMoveSuperimposed();

		//movement done
		IF fbMoveSuperimposed.Done
		THEN
			fbMoveSuperimposed( Execute := FALSE );
			q_xCorrectionActive	:= FALSE;

			SetDiagOutput(	i_etDiag	:= GD.ET_Diag.Ok,
							i_etDiagExt := PDL_ET_DiagExt.WaitForStart,
							i_sMsg		:= '');
			diState	:= 10;

		//user interrupt -> stop and go back to waiting
		ELSIF NOT i_xStart THEN
			fbMoveSuperimposed( Execute := FALSE );
			fbHalt( Execute := FALSE );
			fbHalt(	Axis			:= ifOffsetChannel,
					Execute			:= TRUE,
					BufferMode		:= PLCO.MC_Buffer_Mode.Aborting,
					Deceleration	:= lrCorrAcc );

			q_xCorrectionActive	:= FALSE;
			IF fbHalt.Error THEN
				SetDiagOutput(	i_etDiag	:= GD.ET_Diag.UnexpectedProgramBehavior,
								i_etDiagExt := PDL_ET_DiagExt.UnexpectedFeedback,
								i_sMsg		:= CONCAT('MC_Halt.ErrorId: ', PLCO.FC_EtResultToString(fbHalt.ErrorId) ));
				fbHalt( Execute := FALSE );
				diState := 0;
				RETURN;
			END_IF
			SetDiagOutput(	i_etDiag	:= GD.ET_Diag.Ok,
							i_etDiagExt := PDL_ET_DiagExt.WaitForStart,
							i_sMsg		:= '');
			diState	:= 10;
		END_IF

		//error
		IF fbMoveSuperimposed.Error THEN
			q_xCorrectionActive := FALSE;
			SetDiagOutput(	i_etDiag	:= GD.ET_Diag.UnexpectedProgramBehavior,
							i_etDiagExt := PDL_ET_DiagExt.UnexpectedFeedback,
							i_sMsg		:= CONCAT('MC_MoveSuperimposed.ErrorId: ', TO_STRING(fbMoveSuperimposed.ErrorId)));
			fbMoveSuperimposed( Execute := FALSE );
			diState := 0;
		END_IF
{endregion}

END_CASE

(*--------------------------------------------------------------------------------------------------------------------------------------------*)
